FUNCTION FC 1 : VOID
BEGIN
NETWORK
      A
END_FUNCTION
